(* IEC 61131-3 sources: Aqueous_Solutions/docs-authority/plc (part 4) *)

(* ---- PLC-WTR.st ---- *)
(* AQS-CTL-004 X-CTL-04: control program source, generated by flow_graph/control/plc_programs.py *)
(* Basis: AQS-CTL-001 INSTRUMENT_INDEX.csv, AQS-CTL-002 control architecture, graph set-points. *)
(* PLC-WTR: CPU redundant pair; IO counts AI 71 AO 0 DI 55 DO 10 (modules per AQS-CTL-002, 16-channel, 20 % spare) *)
PROGRAM PLC_WTR_CTRL
VAR
  (* 100 ms cyclic task per AQS-CTL-002 *)
  BMED_UPW_POLISHFT-01_PV : REAL ;  (* S01 normal 2.80 L/h )
  BMED_UPW_POLISHFT-02_PV : REAL ;  (* IA-UPW-FAB normal 2.50 L/h )
  BMED_UPW_POLISHFT-03_PV : REAL ;  (* IA-UPW-REMIN normal 8.98 L/h )
  BMED_UPW_POLISHFT-04_PV : REAL ;  (* IA-UPW-REJ normal 0.25 L/h )
  BMED_UPW_POLISHLT-01_PV : REAL ;  (* A-M-182 liquid height )
  BMED_UPW_POLISHPT-01_PV : REAL ;  (* no design pressure on the graph )
  BMED_UPW_POLISHTE-01_PV : REAL ;  (* band by service )
  CATCH_TANKLT-01_PV : REAL ;  (* A-M-182 liquid height )
  CATCH_TANKPT-01_PV : REAL ;  (* no design pressure on the graph )
  CATCH_TANKTE-01_PV : REAL ;  (* band by service )
  ROOF_TANKFT-01_PV : REAL ;  (* IA-ESS-HYDRO-DIS normal 0.00 L/h )
  ROOF_TANKFT-02_PV : REAL ;  (* S21 normal 5.03 L/h )
  ROOF_TANKFT-03_PV : REAL ;  (* S22 normal 0.00 L/h )
  ROOF_TANKFT-04_PV : REAL ;  (* IA-BED-H2O normal 1.83 L/h )
  ROOF_TANKFT-05_PV : REAL ;  (* IA-DC-SPRAY normal 0.00 L/h )
  ROOF_TANKFT-06_PV : REAL ;  (* IA-NOX-HAB normal 8.64 L/h )
  ROOF_TANKFT-07_PV : REAL ;  (* IA-FLUE-QUENCH normal 1.01 L/h )
  ROOF_TANKFT-08_PV : REAL ;  (* IA-PEROX-H2O normal 0.12 L/h )
  ROOF_TANKFT-09_PV : REAL ;  (* IA-ELY-H2O normal 3.85 L/h )
  ROOF_TANKFT-10_PV : REAL ;  (* IA-CHICK-H2O normal 0.01 L/h )
  ROOF_TANKFT-11_PV : REAL ;  (* IA-AQUA-TOPUP normal 1.14 L/h )
  ROOF_TANKFT-12_PV : REAL ;  (* IA-DUCK-H2O normal 0.08 L/h )
  ROOF_TANKFT-13_PV : REAL ;  (* IA-WASH-FEED normal 0.00 L/h )
  ROOF_TANKFT-14_PV : REAL ;  (* QUAIL_H2O normal 0.01 L/h )
  ROOF_TANKLT-01_PV : REAL ;  (* A-M-182 liquid height )
  ROOF_TANKPT-01_PV : REAL ;  (* no design pressure on the graph )
  ROOF_TANKTE-01_PV : REAL ;  (* band by service )
  BLACK_DIGESTLT-01_PV : REAL ;  (* A-M-182 liquid height )
  BLACK_DIGESTPT-01_PV : REAL ;  (* no design pressure on the graph )
  BLACK_DIGESTTE-01_PV : REAL ;  (* design T 55 C )
  REMINFT-01_PV : REAL ;  (* S26 normal 0.42 L/h )
  REMINFT-02_PV : REAL ;  (* IA-POT-01 normal 8.57 L/h )
  REMINLT-01_PV : REAL ;  (* A-M-182 liquid height )
  REMINPT-01_PV : REAL ;  (* no design pressure on the graph )
  REMINTE-01_PV : REAL ;  (* band by service )
  VCD_TRAINFT-01_PV : REAL ;  (* S25 normal 14.54 L/h )
  VCD_TRAINFT-02_PV : REAL ;  (* S28 normal 0.74 L/h )
  VCD_TRAINFT-03_PV : REAL ;  (* IA-VCD-BD normal 0.28 L/h )
  VCD_TRAINLT-01_PV : REAL ;  (* A-M-182 liquid height )
  VCD_TRAINPT-01_PV : REAL ;  (* no design pressure on the graph )
  VCD_TRAINTE-01_PV : REAL ;  (* band by service )
  GW_INTAKEFT-01_PV : REAL ;  (* IA-GW-MAKEUP normal 0.00 L/h )
  GW_INTAKEFT-02_PV : REAL ;  (* IA-PCA-H2O normal 0.00 L/h )
  GW_INTAKEPT-01_PV : REAL ;  (* no design pressure on the graph )
  GW_INTAKETE-01_PV : REAL ;  (* band by service )
  GREY_TREATFT-01_PV : REAL ;  (* S29 normal 4.35 L/h )
  GREY_TREATFT-02_PV : REAL ;  (* IA-GREY-01 normal 10.75 L/h )
  GREY_TREATFT-03_PV : REAL ;  (* IA-GREY-RET normal 0.00 L/h )
  GREY_TREATLT-01_PV : REAL ;  (* A-M-182 liquid height )
  GREY_TREATPT-01_PV : REAL ;  (* no design pressure on the graph )
  GREY_TREATTE-01_PV : REAL ;  (* band by service )
  GW_INTAKECT-01_PV : REAL ;  (* RO product quality watch; well water moderately mineralised with high silica, fl )
  HDR_UPWPT-01_PV : REAL ;  (* UPW header; no design pressure on the graph )
  HDR_UPWFT-01_PV : REAL ;  (* UPW supply: S01 67.30 kg/d (2.80 L/h) )
  SW_INTAKEFT-01_PV : REAL ;  (* intake delivery watch against the desalination and rejection demand (X-LOC-11 pl )
  DESAL_ROAN-01_PV : REAL ;  (* permeate quality watch against the UPW feed spec (X-LOC-11 placeholder; A-M-410) )
  BRIN_RECOVERAE-01_PV : REAL ;  (* brine concentration watch on the recovery path (X-LOC-11 placeholder; A-M-411) )
  ICE_EXTRACTFT-01_PV : REAL ;  (* melt-water delivery watch against the make-up demand (X-LOC-09 placeholder; A-M- )
  PERC_REMOVEAE-01_PV : REAL ;  (* bed breakthrough watch on the ClO4 reduction (X-LOC-09 placeholder; A-M-407) )
  WET_OXTE-01_PV : REAL ;  (* reactor temperature watch on the wet-oxidation window (X-LOC-10 placeholder; A-M )
  MEM_DISTTE-01_PV : REAL ;  (* feed-permeate temperature difference watch on the membrane loop (X-LOC-10 placeh )
  TANK_BLDPT-01_PV : REAL ;  (* bladder pad pressure gives the water level in the closed tank (X-LOC-09 placehol )
  LB_INTAKEFT-01_PV : REAL ;  (* feed throughput watch against the design 1,000 m3/d (X-LOC-05 Lake Boehmer; A-M- )
  LB_DEGASPT-01_PV : REAL ;  (* air-stripper blower discharge pressure watch at the packing air-to-water ratio ( )
  LB_DEGAS_SCRUBAT-01_PV : REAL ;  (* scrubbed-vent H2S watch against the 10 ppm OSHA ceiling; lethal-site alarm (X-LO )
  LB_SOFTENAT-01_PV : REAL ;  (* lime/soda dosing control on the softened-brine pH (X-LOC-05 Lake Boehmer; A-M-44 )
  LB_ED1PT-01_PV : REAL ;  (* primary ED stack feed pressure watch (X-LOC-05 Lake Boehmer; A-M-438) )
  LB_ED2AT-01_PV : REAL ;  (* product TDS watch against the segment 2311 target (X-LOC-05 Lake Boehmer; A-M-44 )
  LB_PROD_TANKLT-01_PV : REAL ;  (* product buffer level watch (X-LOC-05 Lake Boehmer; A-M-225 basis) )
  LB_BRINE_RETURNFT-01_PV : REAL ;  (* concentrate return flow watch; with the product flow it closes the site salt bal )
  LB_CHEM_STORELT-01_PV : REAL ;  (* chemical day-tank level watch against the resupply interval (X-LOC-05 Lake Boehm )
END_VAR

  (* FLOW control loop - set-point from the graph basis *)
  BMED_UPW_POLISHFT-01_SP := 2.8 ;  (* graph basis: S01 normal 2.80 L/h )
  FB_PI_BMED_UPW_POLISHFT-01( PV := BMED_UPW_POLISHFT-01_PV, SP := BMED_UPW_POLISHFT-01_SP );  (* PI per AQS-CTL-002; GAIN/KI entered at commissioning from the step test (AQS-COM-001 sec. 3), anti-windup clamp per this FB *)
  BMED_UPW_POLISHFT-01_ALARM_HI := 3.08 ;  (* SP x 1.1 margin, A-M-188 margin class *)
  BMED_UPW_POLISHFT-01_ALARM_LO := 2.52 ;

  (* FLOW control loop - set-point from the graph basis *)
  BMED_UPW_POLISHFT-02_SP := 2.5 ;  (* graph basis: IA-UPW-FAB normal 2.50 L/h )
  FB_PI_BMED_UPW_POLISHFT-02( PV := BMED_UPW_POLISHFT-02_PV, SP := BMED_UPW_POLISHFT-02_SP );  (* PI per AQS-CTL-002; GAIN/KI entered at commissioning from the step test (AQS-COM-001 sec. 3), anti-windup clamp per this FB *)
  BMED_UPW_POLISHFT-02_ALARM_HI := 2.75 ;  (* SP x 1.1 margin, A-M-188 margin class *)
  BMED_UPW_POLISHFT-02_ALARM_LO := 2.25 ;

  (* FLOW control loop - set-point from the graph basis *)
  BMED_UPW_POLISHFT-03_SP := 8.98 ;  (* graph basis: IA-UPW-REMIN normal 8.98 L/h )
  FB_PI_BMED_UPW_POLISHFT-03( PV := BMED_UPW_POLISHFT-03_PV, SP := BMED_UPW_POLISHFT-03_SP );  (* PI per AQS-CTL-002; GAIN/KI entered at commissioning from the step test (AQS-COM-001 sec. 3), anti-windup clamp per this FB *)
  BMED_UPW_POLISHFT-03_ALARM_HI := 9.878000000000002 ;  (* SP x 1.1 margin, A-M-188 margin class *)
  BMED_UPW_POLISHFT-03_ALARM_LO := 8.082 ;

  (* FLOW control loop - set-point from the graph basis *)
  BMED_UPW_POLISHFT-04_SP := 0.25 ;  (* graph basis: IA-UPW-REJ normal 0.25 L/h )
  FB_PI_BMED_UPW_POLISHFT-04( PV := BMED_UPW_POLISHFT-04_PV, SP := BMED_UPW_POLISHFT-04_SP );  (* PI per AQS-CTL-002; GAIN/KI entered at commissioning from the step test (AQS-COM-001 sec. 3), anti-windup clamp per this FB *)
  BMED_UPW_POLISHFT-04_ALARM_HI := 0.275 ;  (* SP x 1.1 margin, A-M-188 margin class *)
  BMED_UPW_POLISHFT-04_ALARM_LO := 0.225 ;

  (* LEVEL monitoring block - indication, no set-point invented )
  FB_AI_BMED_UPW_POLISHLT-01( PV := BMED_UPW_POLISHLT-01_PV );
  BMED_UPW_POLISHLT-01_ALARM_HI := 90.0 ;  (* 90 % of span, registered LSH convention )

  (* PRESSURE monitoring block - indication, no set-point invented )
  FB_AI_BMED_UPW_POLISHPT-01( PV := BMED_UPW_POLISHPT-01_PV );
  BMED_UPW_POLISHPT-01_ALARM_HI := 9.0 ;  (* 90 % of span, registered LSH convention )

  (* TEMPERATURE monitoring block - indication, no set-point invented )
  FB_AI_BMED_UPW_POLISHTE-01( PV := BMED_UPW_POLISHTE-01_PV );
  BMED_UPW_POLISHTE-01_ALARM_HI := 135.0 ;  (* 90 % of span, registered LSH convention )

  (* LEVEL monitoring block - indication, no set-point invented )
  FB_AI_CATCH_TANKLT-01( PV := CATCH_TANKLT-01_PV );
  CATCH_TANKLT-01_ALARM_HI := 90.0 ;  (* 90 % of span, registered LSH convention )

  (* PRESSURE monitoring block - indication, no set-point invented )
  FB_AI_CATCH_TANKPT-01( PV := CATCH_TANKPT-01_PV );
  CATCH_TANKPT-01_ALARM_HI := 9.0 ;  (* 90 % of span, registered LSH convention )

  (* TEMPERATURE monitoring block - indication, no set-point invented )
  FB_AI_CATCH_TANKTE-01( PV := CATCH_TANKTE-01_PV );
  CATCH_TANKTE-01_ALARM_HI := 135.0 ;  (* 90 % of span, registered LSH convention )

  (* FLOW control loop - set-point from the graph basis *)
  ROOF_TANKFT-01_SP := 0.0 ;  (* graph basis: IA-ESS-HYDRO-DIS normal 0.00 L/h )
  FB_PI_ROOF_TANKFT-01( PV := ROOF_TANKFT-01_PV, SP := ROOF_TANKFT-01_SP );  (* PI per AQS-CTL-002; GAIN/KI entered at commissioning from the step test (AQS-COM-001 sec. 3), anti-windup clamp per this FB *)
  ROOF_TANKFT-01_ALARM_HI := 0.0 ;  (* expected-zero state: any positive PV alarms )

  (* FLOW control loop - set-point from the graph basis *)
  ROOF_TANKFT-02_SP := 5.03 ;  (* graph basis: S21 normal 5.03 L/h )
  FB_PI_ROOF_TANKFT-02( PV := ROOF_TANKFT-02_PV, SP := ROOF_TANKFT-02_SP );  (* PI per AQS-CTL-002; GAIN/KI entered at commissioning from the step test (AQS-COM-001 sec. 3), anti-windup clamp per this FB *)
  ROOF_TANKFT-02_ALARM_HI := 5.533 ;  (* SP x 1.1 margin, A-M-188 margin class *)
  ROOF_TANKFT-02_ALARM_LO := 4.527 ;

  (* FLOW control loop - set-point from the graph basis *)
  ROOF_TANKFT-03_SP := 0.0 ;  (* graph basis: S22 normal 0.00 L/h )
  FB_PI_ROOF_TANKFT-03( PV := ROOF_TANKFT-03_PV, SP := ROOF_TANKFT-03_SP );  (* PI per AQS-CTL-002; GAIN/KI entered at commissioning from the step test (AQS-COM-001 sec. 3), anti-windup clamp per this FB *)
  ROOF_TANKFT-03_ALARM_HI := 0.0 ;  (* expected-zero state: any positive PV alarms )

  (* FLOW control loop - set-point from the graph basis *)
  ROOF_TANKFT-04_SP := 1.83 ;  (* graph basis: IA-BED-H2O normal 1.83 L/h )
  FB_PI_ROOF_TANKFT-04( PV := ROOF_TANKFT-04_PV, SP := ROOF_TANKFT-04_SP );  (* PI per AQS-CTL-002; GAIN/KI entered at commissioning from the step test (AQS-COM-001 sec. 3), anti-windup clamp per this FB *)
  ROOF_TANKFT-04_ALARM_HI := 2.0130000000000003 ;  (* SP x 1.1 margin, A-M-188 margin class *)
  ROOF_TANKFT-04_ALARM_LO := 1.647 ;

  (* FLOW control loop - set-point from the graph basis *)
  ROOF_TANKFT-05_SP := 0.0 ;  (* graph basis: IA-DC-SPRAY normal 0.00 L/h )
  FB_PI_ROOF_TANKFT-05( PV := ROOF_TANKFT-05_PV, SP := ROOF_TANKFT-05_SP );  (* PI per AQS-CTL-002; GAIN/KI entered at commissioning from the step test (AQS-COM-001 sec. 3), anti-windup clamp per this FB *)
  ROOF_TANKFT-05_ALARM_HI := 0.0 ;  (* expected-zero state: any positive PV alarms )

  (* FLOW control loop - set-point from the graph basis *)
  ROOF_TANKFT-06_SP := 8.64 ;  (* graph basis: IA-NOX-HAB normal 8.64 L/h )
  FB_PI_ROOF_TANKFT-06( PV := ROOF_TANKFT-06_PV, SP := ROOF_TANKFT-06_SP );  (* PI per AQS-CTL-002; GAIN/KI entered at commissioning from the step test (AQS-COM-001 sec. 3), anti-windup clamp per this FB *)
  ROOF_TANKFT-06_ALARM_HI := 9.504000000000001 ;  (* SP x 1.1 margin, A-M-188 margin class *)
  ROOF_TANKFT-06_ALARM_LO := 7.776000000000001 ;

  (* FLOW control loop - set-point from the graph basis *)
  ROOF_TANKFT-07_SP := 1.01 ;  (* graph basis: IA-FLUE-QUENCH normal 1.01 L/h )
  FB_PI_ROOF_TANKFT-07( PV := ROOF_TANKFT-07_PV, SP := ROOF_TANKFT-07_SP );  (* PI per AQS-CTL-002; GAIN/KI entered at commissioning from the step test (AQS-COM-001 sec. 3), anti-windup clamp per this FB *)
  ROOF_TANKFT-07_ALARM_HI := 1.1110000000000002 ;  (* SP x 1.1 margin, A-M-188 margin class *)
  ROOF_TANKFT-07_ALARM_LO := 0.909 ;

  (* FLOW control loop - set-point from the graph basis *)
  ROOF_TANKFT-08_SP := 0.12 ;  (* graph basis: IA-PEROX-H2O normal 0.12 L/h )
  FB_PI_ROOF_TANKFT-08( PV := ROOF_TANKFT-08_PV, SP := ROOF_TANKFT-08_SP );  (* PI per AQS-CTL-002; GAIN/KI entered at commissioning from the step test (AQS-COM-001 sec. 3), anti-windup clamp per this FB *)
  ROOF_TANKFT-08_ALARM_HI := 0.132 ;  (* SP x 1.1 margin, A-M-188 margin class *)
  ROOF_TANKFT-08_ALARM_LO := 0.108 ;

  (* FLOW control loop - set-point from the graph basis *)
  ROOF_TANKFT-09_SP := 3.85 ;  (* graph basis: IA-ELY-H2O normal 3.85 L/h )
  FB_PI_ROOF_TANKFT-09( PV := ROOF_TANKFT-09_PV, SP := ROOF_TANKFT-09_SP );  (* PI per AQS-CTL-002; GAIN/KI entered at commissioning from the step test (AQS-COM-001 sec. 3), anti-windup clamp per this FB *)
  ROOF_TANKFT-09_ALARM_HI := 4.235 ;  (* SP x 1.1 margin, A-M-188 margin class *)
  ROOF_TANKFT-09_ALARM_LO := 3.4650000000000003 ;

  (* FLOW control loop - set-point from the graph basis *)
  ROOF_TANKFT-10_SP := 0.01 ;  (* graph basis: IA-CHICK-H2O normal 0.01 L/h )
  FB_PI_ROOF_TANKFT-10( PV := ROOF_TANKFT-10_PV, SP := ROOF_TANKFT-10_SP );  (* PI per AQS-CTL-002; GAIN/KI entered at commissioning from the step test (AQS-COM-001 sec. 3), anti-windup clamp per this FB *)
  ROOF_TANKFT-10_ALARM_HI := 0.011000000000000001 ;  (* SP x 1.1 margin, A-M-188 margin class *)
  ROOF_TANKFT-10_ALARM_LO := 0.009000000000000001 ;

  (* FLOW control loop - set-point from the graph basis *)
  ROOF_TANKFT-11_SP := 1.14 ;  (* graph basis: IA-AQUA-TOPUP normal 1.14 L/h )
  FB_PI_ROOF_TANKFT-11( PV := ROOF_TANKFT-11_PV, SP := ROOF_TANKFT-11_SP );  (* PI per AQS-CTL-002; GAIN/KI entered at commissioning from the step test (AQS-COM-001 sec. 3), anti-windup clamp per this FB *)
  ROOF_TANKFT-11_ALARM_HI := 1.254 ;  (* SP x 1.1 margin, A-M-188 margin class *)
  ROOF_TANKFT-11_ALARM_LO := 1.026 ;

  (* FLOW control loop - set-point from the graph basis *)
  ROOF_TANKFT-12_SP := 0.08 ;  (* graph basis: IA-DUCK-H2O normal 0.08 L/h )
  FB_PI_ROOF_TANKFT-12( PV := ROOF_TANKFT-12_PV, SP := ROOF_TANKFT-12_SP );  (* PI per AQS-CTL-002; GAIN/KI entered at commissioning from the step test (AQS-COM-001 sec. 3), anti-windup clamp per this FB *)
  ROOF_TANKFT-12_ALARM_HI := 0.08800000000000001 ;  (* SP x 1.1 margin, A-M-188 margin class *)
  ROOF_TANKFT-12_ALARM_LO := 0.07200000000000001 ;

  (* FLOW control loop - set-point from the graph basis *)
  ROOF_TANKFT-13_SP := 0.0 ;  (* graph basis: IA-WASH-FEED normal 0.00 L/h )
  FB_PI_ROOF_TANKFT-13( PV := ROOF_TANKFT-13_PV, SP := ROOF_TANKFT-13_SP );  (* PI per AQS-CTL-002; GAIN/KI entered at commissioning from the step test (AQS-COM-001 sec. 3), anti-windup clamp per this FB *)
  ROOF_TANKFT-13_ALARM_HI := 0.0 ;  (* expected-zero state: any positive PV alarms )

  (* FLOW control loop - set-point from the graph basis *)
  ROOF_TANKFT-14_SP := 0.01 ;  (* graph basis: QUAIL_H2O normal 0.01 L/h )
  FB_PI_ROOF_TANKFT-14( PV := ROOF_TANKFT-14_PV, SP := ROOF_TANKFT-14_SP );  (* PI per AQS-CTL-002; GAIN/KI entered at commissioning from the step test (AQS-COM-001 sec. 3), anti-windup clamp per this FB *)
  ROOF_TANKFT-14_ALARM_HI := 0.011000000000000001 ;  (* SP x 1.1 margin, A-M-188 margin class *)
  ROOF_TANKFT-14_ALARM_LO := 0.009000000000000001 ;

  (* LEVEL monitoring block - indication, no set-point invented )
  FB_AI_ROOF_TANKLT-01( PV := ROOF_TANKLT-01_PV );
  ROOF_TANKLT-01_ALARM_HI := 90.0 ;  (* 90 % of span, registered LSH convention )

  (* PRESSURE monitoring block - indication, no set-point invented )
  FB_AI_ROOF_TANKPT-01( PV := ROOF_TANKPT-01_PV );
  ROOF_TANKPT-01_ALARM_HI := 9.0 ;  (* 90 % of span, registered LSH convention )

  (* TEMPERATURE monitoring block - indication, no set-point invented )
  FB_AI_ROOF_TANKTE-01( PV := ROOF_TANKTE-01_PV );
  ROOF_TANKTE-01_ALARM_HI := 135.0 ;  (* 90 % of span, registered LSH convention )

  (* LEVEL monitoring block - indication, no set-point invented )
  FB_AI_BLACK_DIGESTLT-01( PV := BLACK_DIGESTLT-01_PV );
  BLACK_DIGESTLT-01_ALARM_HI := 90.0 ;  (* 90 % of span, registered LSH convention )

  (* PRESSURE monitoring block - indication, no set-point invented )
  FB_AI_BLACK_DIGESTPT-01( PV := BLACK_DIGESTPT-01_PV );
  BLACK_DIGESTPT-01_ALARM_HI := 9.0 ;  (* 90 % of span, registered LSH convention )

  (* TEMPERATURE control loop - set-point from the graph basis *)
  BLACK_DIGESTTE-01_SP := 55.0 ;  (* graph basis: design T 55 C )
  FB_PI_BLACK_DIGESTTE-01( PV := BLACK_DIGESTTE-01_PV, SP := BLACK_DIGESTTE-01_SP );  (* PI per AQS-CTL-002; GAIN/KI entered at commissioning from the step test (AQS-COM-001 sec. 3), anti-windup clamp per this FB *)
  BLACK_DIGESTTE-01_ALARM_HI := 60.50000000000001 ;  (* SP x 1.1 margin, A-M-188 margin class *)
  BLACK_DIGESTTE-01_ALARM_LO := 49.5 ;

  (* FLOW control loop - set-point from the graph basis *)
  REMINFT-01_SP := 0.42 ;  (* graph basis: S26 normal 0.42 L/h )
  FB_PI_REMINFT-01( PV := REMINFT-01_PV, SP := REMINFT-01_SP );  (* PI per AQS-CTL-002; GAIN/KI entered at commissioning from the step test (AQS-COM-001 sec. 3), anti-windup clamp per this FB *)
  REMINFT-01_ALARM_HI := 0.462 ;  (* SP x 1.1 margin, A-M-188 margin class *)
  REMINFT-01_ALARM_LO := 0.378 ;

  (* FLOW control loop - set-point from the graph basis *)
  REMINFT-02_SP := 8.57 ;  (* graph basis: IA-POT-01 normal 8.57 L/h )
  FB_PI_REMINFT-02( PV := REMINFT-02_PV, SP := REMINFT-02_SP );  (* PI per AQS-CTL-002; GAIN/KI entered at commissioning from the step test (AQS-COM-001 sec. 3), anti-windup clamp per this FB *)
  REMINFT-02_ALARM_HI := 9.427000000000001 ;  (* SP x 1.1 margin, A-M-188 margin class *)
  REMINFT-02_ALARM_LO := 7.713 ;

  (* LEVEL monitoring block - indication, no set-point invented )
  FB_AI_REMINLT-01( PV := REMINLT-01_PV );
  REMINLT-01_ALARM_HI := 90.0 ;  (* 90 % of span, registered LSH convention )

  (* PRESSURE monitoring block - indication, no set-point invented )
  FB_AI_REMINPT-01( PV := REMINPT-01_PV );
  REMINPT-01_ALARM_HI := 9.0 ;  (* 90 % of span, registered LSH convention )

  (* TEMPERATURE monitoring block - indication, no set-point invented )
  FB_AI_REMINTE-01( PV := REMINTE-01_PV );
  REMINTE-01_ALARM_HI := 135.0 ;  (* 90 % of span, registered LSH convention )

  (* FLOW control loop - set-point from the graph basis *)
  VCD_TRAINFT-01_SP := 14.54 ;  (* graph basis: S25 normal 14.54 L/h )
  FB_PI_VCD_TRAINFT-01( PV := VCD_TRAINFT-01_PV, SP := VCD_TRAINFT-01_SP );  (* PI per AQS-CTL-002; GAIN/KI entered at commissioning from the step test (AQS-COM-001 sec. 3), anti-windup clamp per this FB *)
  VCD_TRAINFT-01_ALARM_HI := 15.994 ;  (* SP x 1.1 margin, A-M-188 margin class *)
  VCD_TRAINFT-01_ALARM_LO := 13.086 ;

  (* FLOW control loop - set-point from the graph basis *)
  VCD_TRAINFT-02_SP := 0.74 ;  (* graph basis: S28 normal 0.74 L/h )
  FB_PI_VCD_TRAINFT-02( PV := VCD_TRAINFT-02_PV, SP := VCD_TRAINFT-02_SP );  (* PI per AQS-CTL-002; GAIN/KI entered at commissioning from the step test (AQS-COM-001 sec. 3), anti-windup clamp per this FB *)
  VCD_TRAINFT-02_ALARM_HI := 0.8140000000000001 ;  (* SP x 1.1 margin, A-M-188 margin class *)
  VCD_TRAINFT-02_ALARM_LO := 0.666 ;

  (* FLOW control loop - set-point from the graph basis *)
  VCD_TRAINFT-03_SP := 0.28 ;  (* graph basis: IA-VCD-BD normal 0.28 L/h )
  FB_PI_VCD_TRAINFT-03( PV := VCD_TRAINFT-03_PV, SP := VCD_TRAINFT-03_SP );  (* PI per AQS-CTL-002; GAIN/KI entered at commissioning from the step test (AQS-COM-001 sec. 3), anti-windup clamp per this FB *)
  VCD_TRAINFT-03_ALARM_HI := 0.30800000000000005 ;  (* SP x 1.1 margin, A-M-188 margin class *)
  VCD_TRAINFT-03_ALARM_LO := 0.25200000000000006 ;

  (* LEVEL monitoring block - indication, no set-point invented )
  FB_AI_VCD_TRAINLT-01( PV := VCD_TRAINLT-01_PV );
  VCD_TRAINLT-01_ALARM_HI := 90.0 ;  (* 90 % of span, registered LSH convention )

  (* PRESSURE monitoring block - indication, no set-point invented )
  FB_AI_VCD_TRAINPT-01( PV := VCD_TRAINPT-01_PV );
  VCD_TRAINPT-01_ALARM_HI := 9.0 ;  (* 90 % of span, registered LSH convention )

  (* TEMPERATURE monitoring block - indication, no set-point invented )
  FB_AI_VCD_TRAINTE-01( PV := VCD_TRAINTE-01_PV );
  VCD_TRAINTE-01_ALARM_HI := 135.0 ;  (* 90 % of span, registered LSH convention )

  (* FLOW control loop - set-point from the graph basis *)
  GW_INTAKEFT-01_SP := 0.0 ;  (* graph basis: IA-GW-MAKEUP normal 0.00 L/h )
  FB_PI_GW_INTAKEFT-01( PV := GW_INTAKEFT-01_PV, SP := GW_INTAKEFT-01_SP );  (* PI per AQS-CTL-002; GAIN/KI entered at commissioning from the step test (AQS-COM-001 sec. 3), anti-windup clamp per this FB *)
  GW_INTAKEFT-01_ALARM_HI := 0.0 ;  (* expected-zero state: any positive PV alarms )

  (* FLOW control loop - set-point from the graph basis *)
  GW_INTAKEFT-02_SP := 0.0 ;  (* graph basis: IA-PCA-H2O normal 0.00 L/h )
  FB_PI_GW_INTAKEFT-02( PV := GW_INTAKEFT-02_PV, SP := GW_INTAKEFT-02_SP );  (* PI per AQS-CTL-002; GAIN/KI entered at commissioning from the step test (AQS-COM-001 sec. 3), anti-windup clamp per this FB *)
  GW_INTAKEFT-02_ALARM_HI := 0.0 ;  (* expected-zero state: any positive PV alarms )

  (* PRESSURE monitoring block - indication, no set-point invented )
  FB_AI_GW_INTAKEPT-01( PV := GW_INTAKEPT-01_PV );
  GW_INTAKEPT-01_ALARM_HI := 9.0 ;  (* 90 % of span, registered LSH convention )

  (* TEMPERATURE monitoring block - indication, no set-point invented )
  FB_AI_GW_INTAKETE-01( PV := GW_INTAKETE-01_PV );
  GW_INTAKETE-01_ALARM_HI := 135.0 ;  (* 90 % of span, registered LSH convention )

  (* FLOW control loop - set-point from the graph basis *)
  GREY_TREATFT-01_SP := 4.35 ;  (* graph basis: S29 normal 4.35 L/h )
  FB_PI_GREY_TREATFT-01( PV := GREY_TREATFT-01_PV, SP := GREY_TREATFT-01_SP );  (* PI per AQS-CTL-002; GAIN/KI entered at commissioning from the step test (AQS-COM-001 sec. 3), anti-windup clamp per this FB *)
  GREY_TREATFT-01_ALARM_HI := 4.785 ;  (* SP x 1.1 margin, A-M-188 margin class *)
  GREY_TREATFT-01_ALARM_LO := 3.9149999999999996 ;

  (* FLOW control loop - set-point from the graph basis *)
  GREY_TREATFT-02_SP := 10.75 ;  (* graph basis: IA-GREY-01 normal 10.75 L/h )
  FB_PI_GREY_TREATFT-02( PV := GREY_TREATFT-02_PV, SP := GREY_TREATFT-02_SP );  (* PI per AQS-CTL-002; GAIN/KI entered at commissioning from the step test (AQS-COM-001 sec. 3), anti-windup clamp per this FB *)
  GREY_TREATFT-02_ALARM_HI := 11.825000000000001 ;  (* SP x 1.1 margin, A-M-188 margin class *)
  GREY_TREATFT-02_ALARM_LO := 9.675 ;

  (* FLOW control loop - set-point from the graph basis *)
  GREY_TREATFT-03_SP := 0.0 ;  (* graph basis: IA-GREY-RET normal 0.00 L/h )
  FB_PI_GREY_TREATFT-03( PV := GREY_TREATFT-03_PV, SP := GREY_TREATFT-03_SP );  (* PI per AQS-CTL-002; GAIN/KI entered at commissioning from the step test (AQS-COM-001 sec. 3), anti-windup clamp per this FB *)
  GREY_TREATFT-03_ALARM_HI := 0.0 ;  (* expected-zero state: any positive PV alarms )

  (* LEVEL monitoring block - indication, no set-point invented )
  FB_AI_GREY_TREATLT-01( PV := GREY_TREATLT-01_PV );
  GREY_TREATLT-01_ALARM_HI := 90.0 ;  (* 90 % of span, registered LSH convention )

  (* PRESSURE monitoring block - indication, no set-point invented )
  FB_AI_GREY_TREATPT-01( PV := GREY_TREATPT-01_PV );
  GREY_TREATPT-01_ALARM_HI := 9.0 ;  (* 90 % of span, registered LSH convention )

  (* TEMPERATURE monitoring block - indication, no set-point invented )
  FB_AI_GREY_TREATTE-01( PV := GREY_TREATTE-01_PV );
  GREY_TREATTE-01_ALARM_HI := 135.0 ;  (* 90 % of span, registered LSH convention )

  (* CONDUCTIVITY monitoring block - indication, no set-point invented )
  FB_AI_GW_INTAKECT-01( PV := GW_INTAKECT-01_PV );
  GW_INTAKECT-01_ALARM_HI := 1800.0 ;  (* 90 % of span, registered LSH convention )

  (* PRESSURE monitoring block - indication, no set-point invented )
  FB_AI_HDR_UPWPT-01( PV := HDR_UPWPT-01_PV );
  HDR_UPWPT-01_ALARM_HI := 9.0 ;  (* 90 % of span, registered LSH convention )

  (* FLOW monitoring block - indication, no set-point invented )
  FB_AI_HDR_UPWFT-01( PV := HDR_UPWFT-01_PV );
  HDR_UPWFT-01_ALARM_HI := 9.0 ;  (* 90 % of span, registered LSH convention )

  (* FLOW monitoring block - indication, no set-point invented )
  FB_AI_SW_INTAKEFT-01( PV := SW_INTAKEFT-01_PV );
  SW_INTAKEFT-01_ALARM_HI := 180.0 ;  (* 90 % of span, registered LSH convention )

  (* CONDUCTIVITY monitoring block - indication, no set-point invented )
  FB_AI_DESAL_ROAN-01( PV := DESAL_ROAN-01_PV );
  DESAL_ROAN-01_ALARM_HI := 900.0 ;  (* 90 % of span, registered LSH convention )

  (* COMPOSITION monitoring block - indication, no set-point invented )
  FB_AI_BRIN_RECOVERAE-01( PV := BRIN_RECOVERAE-01_PV );
  BRIN_RECOVERAE-01_ALARM_HI := 135.0 ;  (* 90 % of span, registered LSH convention )

  (* FLOW monitoring block - indication, no set-point invented )
  FB_AI_ICE_EXTRACTFT-01( PV := ICE_EXTRACTFT-01_PV );
  ICE_EXTRACTFT-01_ALARM_HI := 1.8 ;  (* 90 % of span, registered LSH convention )

  (* PERCHLORATE monitoring block - indication, no set-point invented )
  FB_AI_PERC_REMOVEAE-01( PV := PERC_REMOVEAE-01_PV );
  PERC_REMOVEAE-01_ALARM_HI := 90.0 ;  (* 90 % of span, registered LSH convention )

  (* TEMPERATURE monitoring block - indication, no set-point invented )
  FB_AI_WET_OXTE-01( PV := WET_OXTE-01_PV );
  WET_OXTE-01_ALARM_HI := 450.0 ;  (* 90 % of span, registered LSH convention )

  (* TEMPERATURE monitoring block - indication, no set-point invented )
  FB_AI_MEM_DISTTE-01( PV := MEM_DISTTE-01_PV );
  MEM_DISTTE-01_ALARM_HI := 135.0 ;  (* 90 % of span, registered LSH convention )

  (* PRESSURE monitoring block - indication, no set-point invented )
  FB_AI_TANK_BLDPT-01( PV := TANK_BLDPT-01_PV );
  TANK_BLDPT-01_ALARM_HI := 360.0 ;  (* 90 % of span, registered LSH convention )

  (* FLOW monitoring block - indication, no set-point invented )
  FB_AI_LB_INTAKEFT-01( PV := LB_INTAKEFT-01_PV );
  LB_INTAKEFT-01_ALARM_HI := 54.0 ;  (* 90 % of span, registered LSH convention )

  (* PRESSURE monitoring block - indication, no set-point invented )
  FB_AI_LB_DEGASPT-01( PV := LB_DEGASPT-01_PV );
  LB_DEGASPT-01_ALARM_HI := 27.0 ;  (* 90 % of span, registered LSH convention )

  (* HYDROGEN monitoring block - indication, no set-point invented )
  FB_AI_LB_DEGAS_SCRUBAT-01( PV := LB_DEGAS_SCRUBAT-01_PV );
  LB_DEGAS_SCRUBAT-01_ALARM_HI := 45.0 ;  (* 90 % of span, registered LSH convention )

  (* PH monitoring block - indication, no set-point invented )
  FB_AI_LB_SOFTENAT-01( PV := LB_SOFTENAT-01_PV );
  LB_SOFTENAT-01_ALARM_HI := 10.8 ;  (* 90 % of span, registered LSH convention )

  (* PRESSURE monitoring block - indication, no set-point invented )
  FB_AI_LB_ED1PT-01( PV := LB_ED1PT-01_PV );
  LB_ED1PT-01_ALARM_HI := 540.0 ;  (* 90 % of span, registered LSH convention )

  (* CONDUCTIVITY monitoring block - indication, no set-point invented )
  FB_AI_LB_ED2AT-01( PV := LB_ED2AT-01_PV );
  LB_ED2AT-01_ALARM_HI := 27.0 ;  (* 90 % of span, registered LSH convention )

  (* LEVEL monitoring block - indication, no set-point invented )
  FB_AI_LB_PROD_TANKLT-01( PV := LB_PROD_TANKLT-01_PV );
  LB_PROD_TANKLT-01_ALARM_HI := 3.6 ;  (* 90 % of span, registered LSH convention )

  (* FLOW monitoring block - indication, no set-point invented )
  FB_AI_LB_BRINE_RETURNFT-01( PV := LB_BRINE_RETURNFT-01_PV );
  LB_BRINE_RETURNFT-01_ALARM_HI := 36.0 ;  (* 90 % of span, registered LSH convention )

  (* LEVEL monitoring block - indication, no set-point invented )
  FB_AI_LB_CHEM_STORELT-01( PV := LB_CHEM_STORELT-01_PV );
  LB_CHEM_STORELT-01_ALARM_HI := 1.8 ;  (* 90 % of span, registered LSH convention )

END_PROGRAM
